FUNCTION_BLOCK ButtonsPanel (* Composite Function Block Type *)
  (* Standard: 61499-2 *)
  (* Version 0.0, 7/13/2016, Andrei, nxtControl GmbH, template *)
  PACKAGE Main;
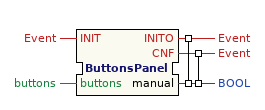
  EVENT_INPUT
    INIT; (* Initialization Request *)
  END_EVENT
  EVENT_OUTPUT
    INITO WITH manual; (* Initialization Confirm *)
    CNF WITH manual;
  END_EVENT
  VAR_OUTPUT
    manual : BOOL;
  END_VAR
  SOCKETS
    buttons : buttons;
  END_SOCKETS
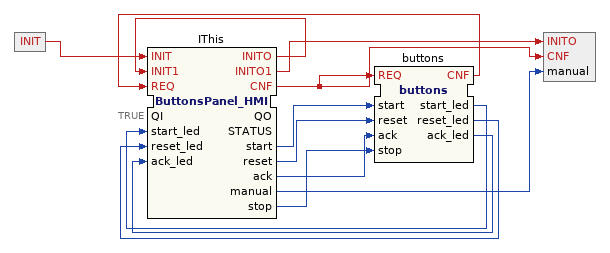
  FBS
    IThis : ButtonsPanel_HMI(QI := TRUE);
  END_FBS
  EVENT_CONNECTIONS
    INIT TO IThis.INIT;
    IThis.INITO TO IThis.INIT1;
    buttons.CNF TO IThis.REQ;
    IThis.INITO1 TO INITO;
    IThis.CNF TO buttons.REQ;
    IThis.CNF TO CNF;
  END_CONNECTIONS
  DATA_CONNECTIONS
    buttons.start_led TO IThis.start_led;
    buttons.reset_led TO IThis.reset_led;
    buttons.ack_led TO IThis.ack_led;
    IThis.start TO buttons.start;
    IThis.reset TO buttons.reset;
    IThis.ack TO buttons.ack;
    IThis.manual TO manual;
    IThis.stop TO buttons.stop;
  END_CONNECTIONS
END_FUNCTION_BLOCK
